Fanuc KAREL source: kb00006.KL

-- PROVISIONAL review KL for V1013-1; original PC SHA256 c23230d1f0108c7e8bd440f2539627c3ad0c14b73dd1147464b360e78e64b794
-- Incomplete behavior may be omitted. Consult companion uncertainty JSON. Do not deploy.
PROGRAM KB00006
%NOLOCKGROUP
BEGIN
  -- UNRESOLVED_PC offsets 5-12; opcodes 9D,23
  -- UNRESOLVED_PC offsets 17-27; opcodes 9D,22,9D,33,35
  -- UNRESOLVED_PC offsets 32-39; opcodes 9D,23
  -- UNRESOLVED_PC offsets 44-51; opcodes 9D,23
  -- UNRESOLVED_PC offsets 56-90; opcodes 27,22,22,22,22,22,31
  -- UNRESOLVED_PC offsets 95-99; opcodes 7F
END KB00006
